(* IEC 61131-3 sources: llm-plc-st-eval/codesys/dobles/A3, 9 files *)

(* ---- 01_Correcta.st ---- *)
(* DOBLE DE PRUEBA A3/Correcta - NO ES CORPUS. Esperado: veredicto 1 *)
FUNCTION_BLOCK FB_Com
VAR_INPUT
    txReq : BOOL;
    rxOk : BOOL;
    rxData : INT;
END_VAR
VAR_OUTPUT
    txData : INT;
    ocupado : BOOL;
    ok : BOOL;
    error : BOOL;
    nIntentos : INT;
END_VAR
VAR
    tPlazo : TON;
    prev : BOOL;
    flanco : BOOL;
END_VAR
flanco := txReq AND NOT prev;
prev := txReq;
IF flanco AND NOT ocupado THEN
    txData := 100;
    ocupado := TRUE;
    ok := FALSE;
    error := FALSE;
    nIntentos := 1;
    tPlazo(IN := FALSE, PT := T#500MS);
ELSIF ocupado THEN
    tPlazo(IN := TRUE, PT := T#500MS);
    IF rxOk AND rxData = txData THEN
        ok := TRUE;
        ocupado := FALSE;
    ELSIF rxOk OR tPlazo.Q THEN
        IF nIntentos < 3 THEN
            nIntentos := nIntentos + 1;
            tPlazo(IN := FALSE, PT := T#500MS);
        ELSE
            error := TRUE;
            ocupado := FALSE;
        END_IF
    END_IF
END_IF
END_FUNCTION_BLOCK

(* ---- 02_PlazoCorto.st ---- *)
(* DOBLE DE PRUEBA A3/PlazoCorto - NO ES CORPUS. Esperado: veredicto 2, falla en el paso 2 *)
FUNCTION_BLOCK FB_Com
VAR_INPUT
    txReq : BOOL;
    rxOk : BOOL;
    rxData : INT;
END_VAR
VAR_OUTPUT
    txData : INT;
    ocupado : BOOL;
    ok : BOOL;
    error : BOOL;
    nIntentos : INT;
END_VAR
VAR
    tPlazo : TON;
    prev : BOOL;
    flanco : BOOL;
END_VAR
flanco := txReq AND NOT prev;
prev := txReq;
IF flanco AND NOT ocupado THEN
    txData := 100;
    ocupado := TRUE;
    ok := FALSE;
    error := FALSE;
    nIntentos := 1;
    tPlazo(IN := FALSE, PT := T#300MS);
ELSIF ocupado THEN
    tPlazo(IN := TRUE, PT := T#300MS);
    IF rxOk AND rxData = txData THEN
        ok := TRUE;
        ocupado := FALSE;
    ELSIF rxOk OR tPlazo.Q THEN
        IF nIntentos < 3 THEN
            nIntentos := nIntentos + 1;
            tPlazo(IN := FALSE, PT := T#300MS);
        ELSE
            error := TRUE;
            ocupado := FALSE;
        END_IF
    END_IF
END_IF
END_FUNCTION_BLOCK

(* ---- 03_PlazoLargo.st ---- *)
(* DOBLE DE PRUEBA A3/PlazoLargo - NO ES CORPUS. Esperado: veredicto 2, falla en el paso 3 *)
FUNCTION_BLOCK FB_Com
VAR_INPUT
    txReq : BOOL;
    rxOk : BOOL;
    rxData : INT;
END_VAR
VAR_OUTPUT
    txData : INT;
    ocupado : BOOL;
    ok : BOOL;
    error : BOOL;
    nIntentos : INT;
END_VAR
VAR
    tPlazo : TON;
    prev : BOOL;
    flanco : BOOL;
END_VAR
flanco := txReq AND NOT prev;
prev := txReq;
IF flanco AND NOT ocupado THEN
    txData := 100;
    ocupado := TRUE;
    ok := FALSE;
    error := FALSE;
    nIntentos := 1;
    tPlazo(IN := FALSE, PT := T#1S);
ELSIF ocupado THEN
    tPlazo(IN := TRUE, PT := T#1S);
    IF rxOk AND rxData = txData THEN
        ok := TRUE;
        ocupado := FALSE;
    ELSIF rxOk OR tPlazo.Q THEN
        IF nIntentos < 3 THEN
            nIntentos := nIntentos + 1;
            tPlazo(IN := FALSE, PT := T#1S);
        ELSE
            error := TRUE;
            ocupado := FALSE;
        END_IF
    END_IF
END_IF
END_FUNCTION_BLOCK

(* ---- 04_PlazoNoSeReinicia.st ---- *)
(* DOBLE DE PRUEBA A3/PlazoNoSeReinicia - NO ES CORPUS. Esperado: veredicto 2, falla en el paso 3 *)
FUNCTION_BLOCK FB_Com
VAR_INPUT
    txReq : BOOL;
    rxOk : BOOL;
    rxData : INT;
END_VAR
VAR_OUTPUT
    txData : INT;
    ocupado : BOOL;
    ok : BOOL;
    error : BOOL;
    nIntentos : INT;
END_VAR
VAR
    tPlazo : TON;
    prev : BOOL;
    flanco : BOOL;
END_VAR
flanco := txReq AND NOT prev;
prev := txReq;
IF flanco AND NOT ocupado THEN
    txData := 100;
    ocupado := TRUE;
    ok := FALSE;
    error := FALSE;
    nIntentos := 1;
    tPlazo(IN := FALSE, PT := T#500MS);
ELSIF ocupado THEN
    tPlazo(IN := TRUE, PT := T#500MS);
    IF rxOk AND rxData = txData THEN
        ok := TRUE;
        ocupado := FALSE;
    ELSIF rxOk OR tPlazo.Q THEN
        IF nIntentos < 3 THEN
            nIntentos := nIntentos + 1;
        ELSE
            error := TRUE;
            ocupado := FALSE;
        END_IF
    END_IF
END_IF
END_FUNCTION_BLOCK

(* ---- 05_IntentosSeBorran.st ---- *)
(* DOBLE DE PRUEBA A3/IntentosSeBorran - NO ES CORPUS. Esperado: veredicto 2, falla en el paso 4 *)
FUNCTION_BLOCK FB_Com
VAR_INPUT
    txReq : BOOL;
    rxOk : BOOL;
    rxData : INT;
END_VAR
VAR_OUTPUT
    txData : INT;
    ocupado : BOOL;
    ok : BOOL;
    error : BOOL;
    nIntentos : INT;
END_VAR
VAR
    tPlazo : TON;
    prev : BOOL;
    flanco : BOOL;
END_VAR
flanco := txReq AND NOT prev;
prev := txReq;
IF flanco AND NOT ocupado THEN
    txData := 100;
    ocupado := TRUE;
    ok := FALSE;
    error := FALSE;
    nIntentos := 1;
    tPlazo(IN := FALSE, PT := T#500MS);
ELSIF ocupado THEN
    tPlazo(IN := TRUE, PT := T#500MS);
    IF rxOk AND rxData = txData THEN
        ok := TRUE;
        ocupado := FALSE;
    ELSIF rxOk OR tPlazo.Q THEN
        IF nIntentos < 3 THEN
            nIntentos := nIntentos + 1;
            tPlazo(IN := FALSE, PT := T#500MS);
        ELSE
            error := TRUE;
            ocupado := FALSE;
        END_IF
    END_IF
END_IF
IF NOT ocupado THEN
    nIntentos := 0;
END_IF
END_FUNCTION_BLOCK

(* ---- 06_OkNoSeBorra.st ---- *)
(* DOBLE DE PRUEBA A3/OkNoSeBorra - NO ES CORPUS. Esperado: veredicto 2, falla en el paso 6 *)
FUNCTION_BLOCK FB_Com
VAR_INPUT
    txReq : BOOL;
    rxOk : BOOL;
    rxData : INT;
END_VAR
VAR_OUTPUT
    txData : INT;
    ocupado : BOOL;
    ok : BOOL;
    error : BOOL;
    nIntentos : INT;
END_VAR
VAR
    tPlazo : TON;
    prev : BOOL;
    flanco : BOOL;
END_VAR
flanco := txReq AND NOT prev;
prev := txReq;
IF flanco AND NOT ocupado THEN
    txData := 100;
    ocupado := TRUE;
    nIntentos := 1;
    tPlazo(IN := FALSE, PT := T#500MS);
ELSIF ocupado THEN
    tPlazo(IN := TRUE, PT := T#500MS);
    IF rxOk AND rxData = txData THEN
        ok := TRUE;
        ocupado := FALSE;
    ELSIF rxOk OR tPlazo.Q THEN
        IF nIntentos < 3 THEN
            nIntentos := nIntentos + 1;
            tPlazo(IN := FALSE, PT := T#500MS);
        ELSE
            error := TRUE;
            ocupado := FALSE;
        END_IF
    END_IF
END_IF
END_FUNCTION_BLOCK

(* ---- 07_SinEco.st ---- *)
(* DOBLE DE PRUEBA A3/SinEco - NO ES CORPUS. Esperado: veredicto 2, falla en el paso 7 *)
FUNCTION_BLOCK FB_Com
VAR_INPUT
    txReq : BOOL;
    rxOk : BOOL;
    rxData : INT;
END_VAR
VAR_OUTPUT
    txData : INT;
    ocupado : BOOL;
    ok : BOOL;
    error : BOOL;
    nIntentos : INT;
END_VAR
VAR
    tPlazo : TON;
    prev : BOOL;
    flanco : BOOL;
END_VAR
flanco := txReq AND NOT prev;
prev := txReq;
IF flanco AND NOT ocupado THEN
    txData := 100;
    ocupado := TRUE;
    ok := FALSE;
    error := FALSE;
    nIntentos := 1;
    tPlazo(IN := FALSE, PT := T#500MS);
ELSIF ocupado THEN
    tPlazo(IN := TRUE, PT := T#500MS);
    IF rxOk THEN
        ok := TRUE;
        ocupado := FALSE;
    ELSIF rxOk OR tPlazo.Q THEN
        IF nIntentos < 3 THEN
            nIntentos := nIntentos + 1;
            tPlazo(IN := FALSE, PT := T#500MS);
        ELSE
            error := TRUE;
            ocupado := FALSE;
        END_IF
    END_IF
END_IF
END_FUNCTION_BLOCK

(* ---- 08_ReiniciaPorTxReq.st ---- *)
(* DOBLE DE PRUEBA A3/ReiniciaPorTxReq - NO ES CORPUS. Esperado: veredicto 2, falla en el paso 8 *)
FUNCTION_BLOCK FB_Com
VAR_INPUT
    txReq : BOOL;
    rxOk : BOOL;
    rxData : INT;
END_VAR
VAR_OUTPUT
    txData : INT;
    ocupado : BOOL;
    ok : BOOL;
    error : BOOL;
    nIntentos : INT;
END_VAR
VAR
    tPlazo : TON;
    prev : BOOL;
    flanco : BOOL;
END_VAR
flanco := txReq AND NOT prev;
prev := txReq;
IF flanco THEN
    txData := 100;
    ocupado := TRUE;
    ok := FALSE;
    error := FALSE;
    nIntentos := 1;
    tPlazo(IN := FALSE, PT := T#500MS);
ELSIF ocupado THEN
    tPlazo(IN := TRUE, PT := T#500MS);
    IF rxOk AND rxData = txData THEN
        ok := TRUE;
        ocupado := FALSE;
    ELSIF rxOk OR tPlazo.Q THEN
        IF nIntentos < 3 THEN
            nIntentos := nIntentos + 1;
            tPlazo(IN := FALSE, PT := T#500MS);
        ELSE
            error := TRUE;
            ocupado := FALSE;
        END_IF
    END_IF
END_IF
END_FUNCTION_BLOCK

(* ---- 09_CuatroIntentos.st ---- *)
(* DOBLE DE PRUEBA A3/CuatroIntentos - NO ES CORPUS. Esperado: veredicto 2, falla en el paso 10 *)
FUNCTION_BLOCK FB_Com
VAR_INPUT
    txReq : BOOL;
    rxOk : BOOL;
    rxData : INT;
END_VAR
VAR_OUTPUT
    txData : INT;
    ocupado : BOOL;
    ok : BOOL;
    error : BOOL;
    nIntentos : INT;
END_VAR
VAR
    tPlazo : TON;
    prev : BOOL;
    flanco : BOOL;
END_VAR
flanco := txReq AND NOT prev;
prev := txReq;
IF flanco AND NOT ocupado THEN
    txData := 100;
    ocupado := TRUE;
    ok := FALSE;
    error := FALSE;
    nIntentos := 1;
    tPlazo(IN := FALSE, PT := T#500MS);
ELSIF ocupado THEN
    tPlazo(IN := TRUE, PT := T#500MS);
    IF rxOk AND rxData = txData THEN
        ok := TRUE;
        ocupado := FALSE;
    ELSIF rxOk OR tPlazo.Q THEN
        IF nIntentos < 4 THEN
            nIntentos := nIntentos + 1;
            tPlazo(IN := FALSE, PT := T#500MS);
        ELSE
            error := TRUE;
            ocupado := FALSE;
        END_IF
    END_IF
END_IF
END_FUNCTION_BLOCK
